// Mitsubishi GX Works2 project: Bloque A   PLC: FX2N/FX2NC

PROGRAM MAIN
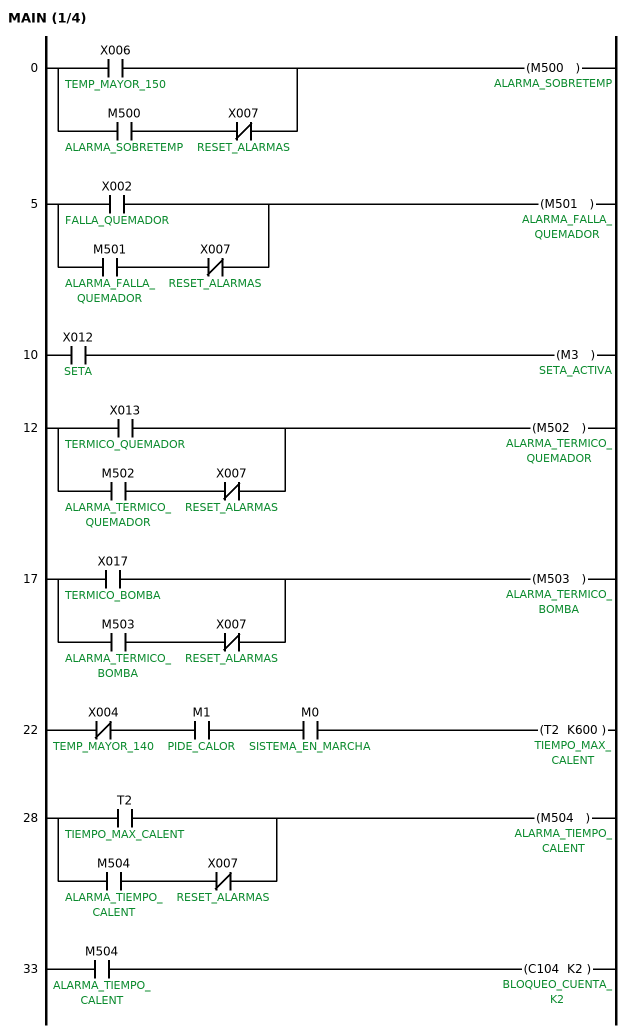
0     LD      X006  ; TEMP_MAYOR_150
      LD      M500  ; ALARMA_SOBRETEMP
      ANI     X007  ; RESET_ALARMAS
      ORB
      OUT     M500  ; ALARMA_SOBRETEMP
5     LD      X002  ; FALLA_QUEMADOR
      LD      M501  ; ALARMA_FALLA_QUEMADOR
      ANI     X007  ; RESET_ALARMAS
      ORB
      OUT     M501  ; ALARMA_FALLA_QUEMADOR
10    LD      X012  ; SETA
      OUT     M3  ; SETA_ACTIVA
12    LD      X013  ; TERMICO_QUEMADOR
      LD      M502  ; ALARMA_TERMICO_QUEMADOR
      ANI     X007  ; RESET_ALARMAS
      ORB
      OUT     M502  ; ALARMA_TERMICO_QUEMADOR
17    LD      X017  ; TERMICO_BOMBA
      LD      M503  ; ALARMA_TERMICO_BOMBA
      ANI     X007  ; RESET_ALARMAS
      ORB
      OUT     M503  ; ALARMA_TERMICO_BOMBA
22    LDI     X004  ; TEMP_MAYOR_140
      AND     M1  ; PIDE_CALOR
      AND     M0  ; SISTEMA_EN_MARCHA
      OUT     T2 K600  ; TIEMPO_MAX_CALENT
28    LD      T2  ; TIEMPO_MAX_CALENT
      LD      M504  ; ALARMA_TIEMPO_CALENT
      ANI     X007  ; RESET_ALARMAS
      ORB
      OUT     M504  ; ALARMA_TIEMPO_CALENT
33    LD      M504  ; ALARMA_TIEMPO_CALENT
      OUT     C104 K2  ; BLOQUEO_CUENTA_K2
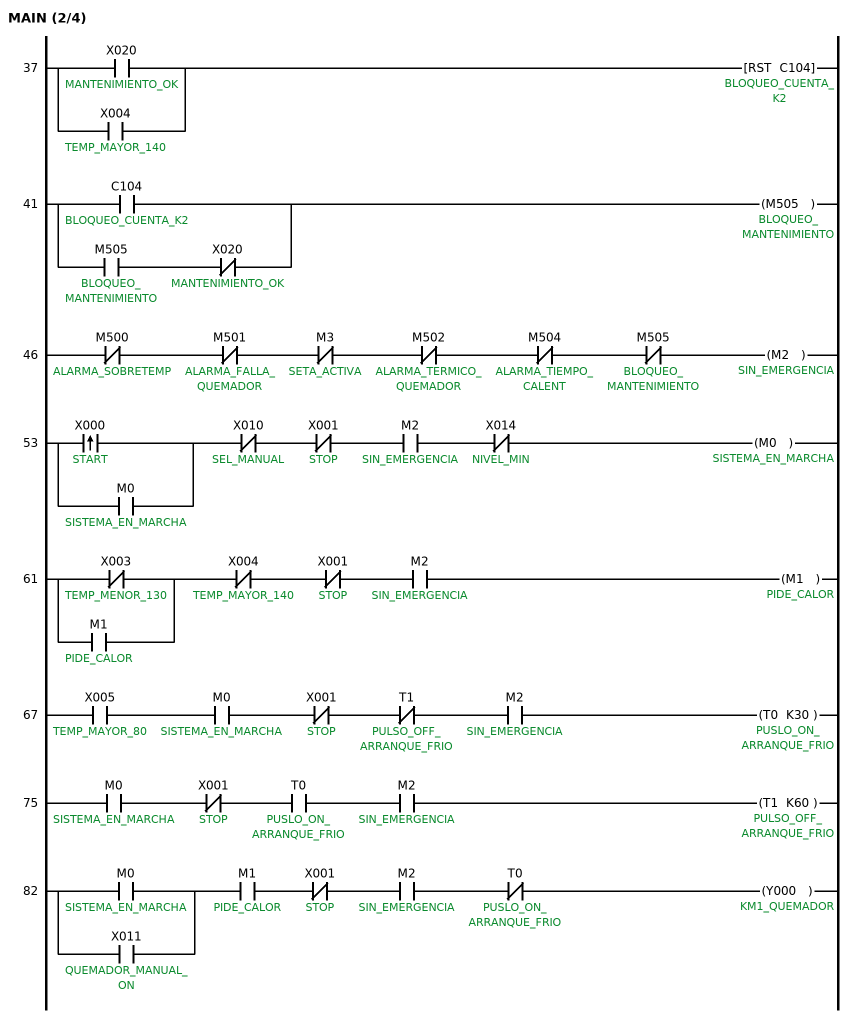
37    LD      X020  ; MANTENIMIENTO_OK
      OR      X004  ; TEMP_MAYOR_140
      RST     C104  ; BLOQUEO_CUENTA_K2
41    LD      C104  ; BLOQUEO_CUENTA_K2
      LD      M505  ; BLOQUEO_MANTENIMIENTO
      ANI     X020  ; MANTENIMIENTO_OK
      ORB
      OUT     M505  ; BLOQUEO_MANTENIMIENTO
46    LDI     M500  ; ALARMA_SOBRETEMP
      ANI     M501  ; ALARMA_FALLA_QUEMADOR
      ANI     M3  ; SETA_ACTIVA
      ANI     M502  ; ALARMA_TERMICO_QUEMADOR
      ANI     M504  ; ALARMA_TIEMPO_CALENT
      ANI     M505  ; BLOQUEO_MANTENIMIENTO
      OUT     M2  ; SIN_EMERGENCIA
53    LDP     X000  ; START
      OR      M0  ; SISTEMA_EN_MARCHA
      ANI     X010  ; SEL_MANUAL
      ANI     X001  ; STOP
      AND     M2  ; SIN_EMERGENCIA
      ANI     X014  ; NIVEL_MIN
      OUT     M0  ; SISTEMA_EN_MARCHA
61    LDI     X003  ; TEMP_MENOR_130
      OR      M1  ; PIDE_CALOR
      ANI     X004  ; TEMP_MAYOR_140
      ANI     X001  ; STOP
      AND     M2  ; SIN_EMERGENCIA
      OUT     M1  ; PIDE_CALOR
67    LD      X005  ; TEMP_MAYOR_80
      AND     M0  ; SISTEMA_EN_MARCHA
      ANI     X001  ; STOP
      ANI     T1  ; PULSO_OFF_ARRANQUE_FRIO
      AND     M2  ; SIN_EMERGENCIA
      OUT     T0 K30  ; PUSLO_ON_ARRANQUE_FRIO
75    LD      M0  ; SISTEMA_EN_MARCHA
      ANI     X001  ; STOP
      AND     T0  ; PUSLO_ON_ARRANQUE_FRIO
      AND     M2  ; SIN_EMERGENCIA
      OUT     T1 K60  ; PULSO_OFF_ARRANQUE_FRIO
82    LD      M0  ; SISTEMA_EN_MARCHA
      OR      X011  ; QUEMADOR_MANUAL_ON
      AND     M1  ; PIDE_CALOR
      ANI     X001  ; STOP
      AND     M2  ; SIN_EMERGENCIA
      ANI     T0  ; PUSLO_ON_ARRANQUE_FRIO
      OUT     Y000  ; KM1_QUEMADOR
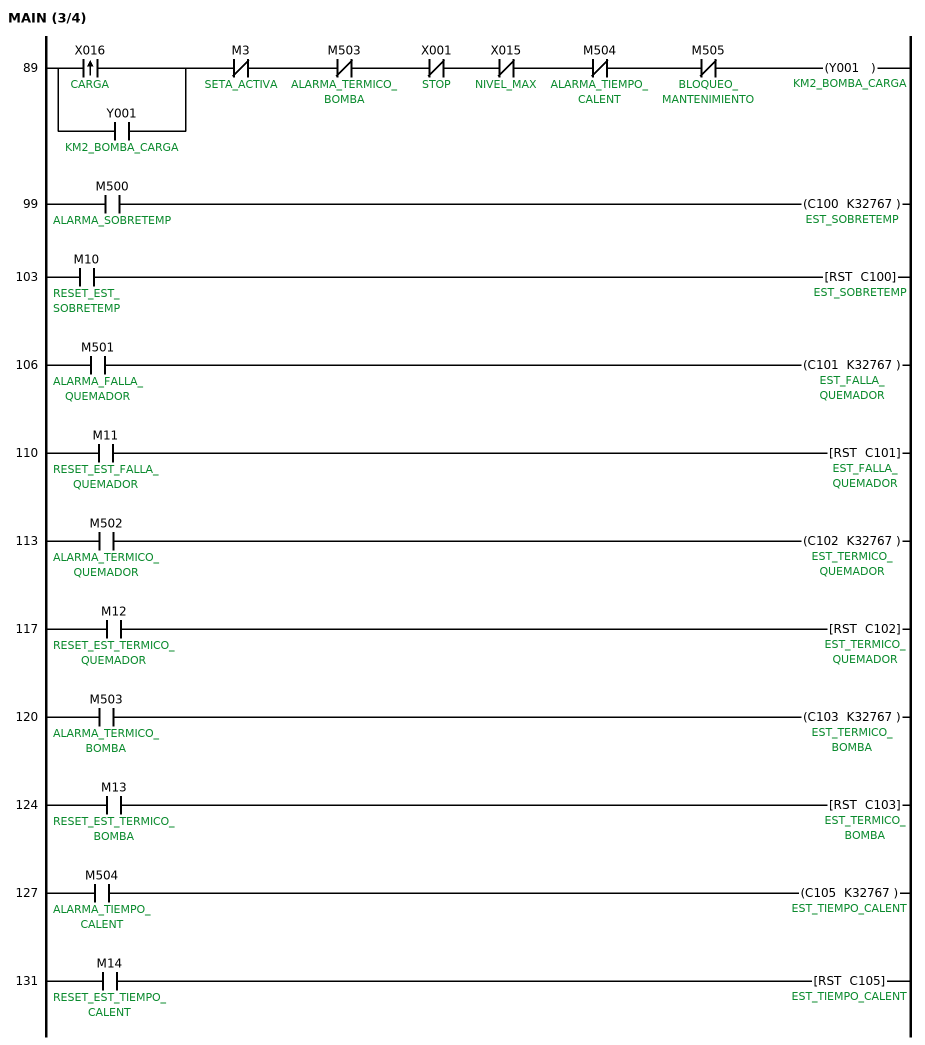
89    LDP     X016  ; CARGA
      OR      Y001  ; KM2_BOMBA_CARGA
      ANI     M3  ; SETA_ACTIVA
      ANI     M503  ; ALARMA_TERMICO_BOMBA
      ANI     X001  ; STOP
      ANI     X015  ; NIVEL_MAX
      ANI     M504  ; ALARMA_TIEMPO_CALENT
      ANI     M505  ; BLOQUEO_MANTENIMIENTO
      OUT     Y001  ; KM2_BOMBA_CARGA
99    LD      M500  ; ALARMA_SOBRETEMP
      OUT     C100 K32767  ; EST_SOBRETEMP
103   LD      M10  ; RESET_EST_SOBRETEMP
      RST     C100  ; EST_SOBRETEMP
106   LD      M501  ; ALARMA_FALLA_QUEMADOR
      OUT     C101 K32767  ; EST_FALLA_QUEMADOR
110   LD      M11  ; RESET_EST_FALLA_QUEMADOR
      RST     C101  ; EST_FALLA_QUEMADOR
113   LD      M502  ; ALARMA_TERMICO_QUEMADOR
      OUT     C102 K32767  ; EST_TERMICO_QUEMADOR
117   LD      M12  ; RESET_EST_TERMICO_QUEMADOR
      RST     C102  ; EST_TERMICO_QUEMADOR
120   LD      M503  ; ALARMA_TERMICO_BOMBA
      OUT     C103 K32767  ; EST_TERMICO_BOMBA
124   LD      M13  ; RESET_EST_TERMICO_BOMBA
      RST     C103  ; EST_TERMICO_BOMBA
127   LD      M504  ; ALARMA_TIEMPO_CALENT
      OUT     C105 K32767  ; EST_TIEMPO_CALENT
131   LD      M14  ; RESET_EST_TIEMPO_CALENT
      RST     C105  ; EST_TIEMPO_CALENT
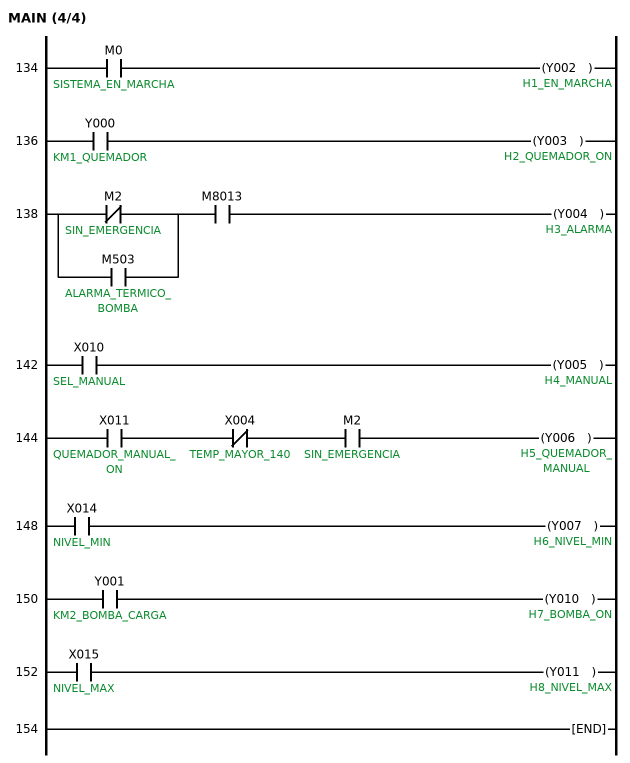
134   LD      M0  ; SISTEMA_EN_MARCHA
      OUT     Y002  ; H1_EN_MARCHA
136   LD      Y000  ; KM1_QUEMADOR
      OUT     Y003  ; H2_QUEMADOR_ON
138   LDI     M2  ; SIN_EMERGENCIA
      OR      M503  ; ALARMA_TERMICO_BOMBA
      AND     M8013
      OUT     Y004  ; H3_ALARMA
142   LD      X010  ; SEL_MANUAL
      OUT     Y005  ; H4_MANUAL
144   LD      X011  ; QUEMADOR_MANUAL_ON
      ANI     X004  ; TEMP_MAYOR_140
      AND     M2  ; SIN_EMERGENCIA
      OUT     Y006  ; H5_QUEMADOR_MANUAL
148   LD      X014  ; NIVEL_MIN
      OUT     Y007  ; H6_NIVEL_MIN
150   LD      Y001  ; KM2_BOMBA_CARGA
      OUT     Y010  ; H7_BOMBA_ON
152   LD      X015  ; NIVEL_MAX
      OUT     Y011  ; H8_NIVEL_MAX
154   END
END_PROGRAM
